TYPE SimulatorFeedback :
STRUCT
	version : UDINT;
	sequence : UDINT;
	timeInNs : ULINT;
	leftWheelAngleInRad : LREAL;
	rightWheelAngleInRad : LREAL;
	leftWheelVelocityInRadPerS : LREAL;
	rightWheelVelocityInRadPerS : LREAL;
	angularRateInRadPerS : Vector3;
	accelerationInMPerS2 : Vector3;
	truePose : Pose2D;
	collided : BOOL;
END_STRUCT
END_TYPE

(* stored: Version 1.1.0.1, ProductVersion 3.1.4026.12
   DUT SimulatorFeedback: Id {e9abb3ad-d5f3-5e82-9664-324ad1e56666} *)
